Staubli VAL3: toolItem.pjx

--- toolItem.pjx ---
Parameters version=s8.10.3Cs9_BS2093 stackSize=5000 millimeterUnit=true
Program file=start.pgx
Program file=stop.pgx
Data file=toolItem.dtx

--- toolItem.dtx ---
public string sName
public tool tTool = {fatherId=flange[0]}

--- start.pgx ---
program start()
begin
end

--- stop.pgx ---
program stop()
begin
end
